(* IEC 61131-3 sources: stdmachine/plc/src/03_Base, 34 files *)

(* ---- GVL_BeaconBits.st ---- *)
// Codage de la balise (ST_MachineStatus.nBeacon, ST_StationStatus.nBeacon, I_Beacon.SetPattern)
{attribute 'qualified_only'}
VAR_GLOBAL CONSTANT
    RED : UINT := 16#0001;
    ORANGE : UINT := 16#0002;
    GREEN : UINT := 16#0004;
    BLUE : UINT := 16#0008;
    RED_BLINK : UINT := 16#0100;
    ORANGE_BLINK : UINT := 16#0200;
    GREEN_BLINK : UINT := 16#0400;
    BLUE_BLINK : UINT := 16#0800;
    BUZZER : UINT := 16#1000;
END_VAR

(* ---- GVL_Curves.st ---- *)
// Courbes de presse (docs/05 § 9) : tampon circulaire GVL_Hmi.aCurve[1..8], dernière courbe de chaque station
// pour la trace de l'opération (ST_TraceRecord.nCurveId).
{attribute 'qualified_only'}
VAR_GLOBAL
    nNextCurveId : UDINT := 1;
    nNextSlot : USINT := 1;
    aLastCurveId : ARRAY[0..GVL_Const.MAX_STATIONS] OF UDINT;
    aLastCurveTime : ARRAY[0..GVL_Const.MAX_STATIONS] OF LINT;      // début de l'enregistrement (UTC)
END_VAR

(* ---- GVL_IoRef.st ---- *)
// Pointeurs vers l'image E/S et les pools matériels du projet de la machine (docs/04 § 6).
// GVL_IO et GVL_Hw sont dans le projet de la machine (reliés aux bornes) ; MAIN les donne ici au premier cycle :
//     GVL_IoRef.pDI := ADR(GVL_IO.aDI); … ; GVL_IoRef.pAxis := ADR(GVL_Hw.aAxis); GVL_IoRef.nAxes := …
{attribute 'qualified_only'}
VAR_GLOBAL
    pDI : POINTER TO ARRAY[0..GVL_Const.MAX_DI - 1] OF BOOL;
    pDO : POINTER TO ARRAY[0..GVL_Const.MAX_DO - 1] OF BOOL;
    pAI : POINTER TO ARRAY[0..GVL_Const.MAX_AI - 1] OF INT;
    pAO : POINTER TO ARRAY[0..GVL_Const.MAX_AO - 1] OF INT;
    pAxis : POINTER TO ARRAY[1..GVL_Const.MAX_AXES] OF AXIS_REF;   // GVL_Hw.aAxis
    nAxes : INT;                     // nombre d'axes reliés dans GVL_Hw
    // Rempli par FB_Machine au premier cycle, pour les objets Système planaire et Mover
    ipPlanar : I_PlanarDriver;
    ipMovers : I_MoverMotion;
END_VAR

(* ---- GVL_Sim.st ---- *)
// Simulation de toute la machine (docs/04 § 6.3)
{attribute 'qualified_only'}
VAR_GLOBAL
    bAllSimulated : BOOL;
    nSeed : UDINT := 16#2545F491;      // générateur pseudo-aléatoire des objets simulés (F_SimRandom)
END_VAR

(* ---- F_AddDeployError.st ---- *)
// Ajoute une erreur à la réponse de déploiement (docs/05 § 10, étape 5) ; les codes sont listés dans FB_Loader
FUNCTION F_AddDeployError : BOOL
VAR_IN_OUT
    stResp : ST_DeployResponse;
END_VAR
VAR_INPUT
    nCode : UINT;
    nStation : USINT;
    nTable : USINT;
    nInstr : INT;
    nObject : UINT;
    nDetail : UDINT;
END_VAR
F_AddDeployError := FALSE;
IF stResp.nErrors >= 32 THEN RETURN; END_IF       // les suivantes sont perdues : 32 suffisent pour corriger
stResp.nErrors := stResp.nErrors + 1;
stResp.aError[stResp.nErrors].nCode := nCode;
stResp.aError[stResp.nErrors].nStation := nStation;
stResp.aError[stResp.nErrors].nTable := nTable;
stResp.aError[stResp.nErrors].nInstr := nInstr;
stResp.aError[stResp.nErrors].nObject := nObject;
stResp.aError[stResp.nErrors].nDetail := nDetail;
F_AddDeployError := TRUE;
END_FUNCTION

(* ---- F_AddRetained.st ---- *)
// Ajoute une valeur à la liste publiée pour la sauvegarde par la HMI (docs/02 § 7.4)
FUNCTION F_AddRetained : BOOL
VAR_IN_OUT
    stOut : ST_RetainedValues;
    stItem : ST_RetainedItem;
END_VAR
F_AddRetained := FALSE;
IF stOut.nCount >= 2048 THEN RETURN; END_IF
stOut.nCount := stOut.nCount + 1;
stOut.aItem[stOut.nCount] := stItem;
F_AddRetained := TRUE;
END_FUNCTION

(* ---- F_AggregateState.st ---- *)
// État agrégé d'un parent : En erreur > Non initialisé > En cours > Prêt (docs/04 § 8)
FUNCTION F_AggregateState : E_ObjState
VAR_INPUT
    eCurrent : E_ObjState;       // agrégat en cours de calcul
    eChild : E_ObjState;
END_VAR
IF eCurrent = E_ObjState.Error OR eChild = E_ObjState.Error THEN
    F_AggregateState := E_ObjState.Error;
ELSIF eCurrent = E_ObjState.NotInitialized OR eChild = E_ObjState.NotInitialized THEN
    F_AggregateState := E_ObjState.NotInitialized;
ELSIF eCurrent = E_ObjState.Busy OR eChild = E_ObjState.Busy THEN
    F_AggregateState := E_ObjState.Busy;
ELSE
    F_AggregateState := E_ObjState.Ready;
END_IF

(* ---- F_ApplyOp.st ---- *)
// SetVar : 0 affecter, 1 ajouter, 2 soustraire (docs/06 § 3)
FUNCTION F_ApplyOp : LREAL
VAR_INPUT
    fCurrent : LREAL;
    fValue : LREAL;
    nOp : DINT;
END_VAR
CASE nOp OF
    1: F_ApplyOp := fCurrent + fValue;
    2: F_ApplyOp := fCurrent - fValue;
ELSE
    F_ApplyOp := fValue;
END_CASE

(* ---- F_AxisRef.st ---- *)
// Pointeur vers l'axe NC n° nDevice du pool matériel (docs/04 § 6.2) ; 0 si absent
FUNCTION F_AxisRef : POINTER TO AXIS_REF
VAR_INPUT
    nDevice : INT;
END_VAR
IF GVL_IoRef.pAxis = 0 OR nDevice < 1 OR nDevice > GVL_IoRef.nAxes OR nDevice > GVL_Const.MAX_AXES THEN
    F_AxisRef := 0;
ELSE
    F_AxisRef := ADR(GVL_IoRef.pAxis^[nDevice]);
END_IF

(* ---- F_BeaconPattern.st ---- *)
// Couleurs de la balise selon l'état (docs/02 § 8, tableau des balises)
FUNCTION F_BeaconPattern : UINT
VAR_INPUT
    eState : E_State;
    bMaintenance : BOOL;         // mode Maintenance, ou état déclaré maintenance, essais, nettoyage
    bOperatorAwaited : BOOL;     // mover à vider, fin d'OF, machine vidée, réaction qualité…
    bStationAborted : BOOL;      // machine : une station Aborted pendant que la machine produit
END_VAR
VAR
    n : UINT;
END_VAR
CASE eState OF
    E_State.Execute:
        n := GVL_BeaconBits.GREEN;
        IF bStationAborted THEN n := n OR GVL_BeaconBits.RED_BLINK; END_IF
    E_State.Idle:
        n := GVL_BeaconBits.GREEN_BLINK;
    E_State.Held, E_State.Stopped:
        n := GVL_BeaconBits.ORANGE;
    E_State.Resetting, E_State.Stopping, E_State.Clearing:
        n := GVL_BeaconBits.ORANGE_BLINK;
    E_State.Aborted:
        n := GVL_BeaconBits.RED_BLINK OR GVL_BeaconBits.BUZZER;
END_CASE
IF bMaintenance THEN n := n OR GVL_BeaconBits.BLUE; END_IF
IF bOperatorAwaited THEN n := n OR GVL_BeaconBits.BLUE_BLINK; END_IF
F_BeaconPattern := n;

(* ---- F_CalibStateNum.st ---- *)
// État de calibration ↔ nombre, pour la sauvegarde des valeurs par la HMI (ST_RetainedItem.aValue[1])
FUNCTION F_CalibStateNum : LREAL
VAR_INPUT
    eState : E_CalibState;
END_VAR
CASE eState OF
    E_CalibState.Valid: F_CalibStateNum := 1;
    E_CalibState.Expired: F_CalibStateNum := 2;
    E_CalibState.Failed: F_CalibStateNum := 3;
    E_CalibState.Running: F_CalibStateNum := 4;
ELSE
    F_CalibStateNum := 0;
END_CASE
END_FUNCTION

(* ---- F_CalibStateOf.st ---- *)
// Nombre → état de calibration (restauration) ; une calibration en cours à la sauvegarde revient « jamais faite »
FUNCTION F_CalibStateOf : E_CalibState
VAR_INPUT
    fValue : LREAL;
END_VAR
IF fValue > 2.5 AND fValue < 3.5 THEN
    F_CalibStateOf := E_CalibState.Failed;
ELSIF fValue > 1.5 AND fValue < 2.5 THEN
    F_CalibStateOf := E_CalibState.Expired;
ELSIF fValue > 0.5 AND fValue < 1.5 THEN
    F_CalibStateOf := E_CalibState.Valid;
ELSE
    F_CalibStateOf := E_CalibState.Never;
END_IF
END_FUNCTION

(* ---- F_CatalogBit.st ---- *)
// Vrai si le bit de l'action est posé dans un masque du catalogue (GVL_Catalog.a*Mask)
FUNCTION F_CatalogBit : BOOL
VAR_INPUT
    nMask : UDINT;
    nAction : UINT;
END_VAR
IF nAction < 1 OR nAction > GVL_Const.MAX_ACTION THEN
    F_CatalogBit := FALSE;
ELSE
    F_CatalogBit := (SHR(nMask, nAction - 1) AND 1) = 1;
END_IF

(* ---- F_CatalogHasAction.st ---- *)
// L'action existe-t-elle pour ce type ? (docs/04 § 7.3)
FUNCTION F_CatalogHasAction : BOOL
VAR_INPUT
    nType : UINT;
    nAction : UINT;
END_VAR
IF nType > GVL_Const.MAX_TYPE THEN
    F_CatalogHasAction := FALSE;
ELSE
    F_CatalogHasAction := F_CatalogBit(GVL_Catalog.aActionMask[nType], nAction);
END_IF

(* ---- F_Compare.st ---- *)
// Terme de condition (docs/05 § 3.7) : égalités sur réels à 1e-9 près
FUNCTION F_Compare : BOOL
VAR_INPUT
    a : LREAL;
    eCmp : E_Cmp;
    b : LREAL;
END_VAR
CASE eCmp OF
    E_Cmp.Eq: F_Compare := ABS(a - b) < 1.0E-9;
    E_Cmp.Ne: F_Compare := ABS(a - b) >= 1.0E-9;
    E_Cmp.Lt: F_Compare := a < b;
    E_Cmp.Le: F_Compare := a <= b + 1.0E-9;
    E_Cmp.Gt: F_Compare := a > b;
    E_Cmp.Ge: F_Compare := a >= b - 1.0E-9;
    E_Cmp.IsTrue: F_Compare := a <> 0;
    E_Cmp.IsFalse: F_Compare := a = 0;
ELSE
    F_Compare := FALSE;
END_CASE

(* ---- F_CycleMs.st ---- *)
// Durée du cycle de la tâche courante en ms (docs/04 § 2)
FUNCTION F_CycleMs : LREAL
VAR
    nTask : DINT;
END_VAR
nTask := GETCURTASKINDEXEX();
F_CycleMs := UDINT_TO_LREAL(TwinCAT_SystemInfoVarList._TaskInfo[nTask].CycleTime) / 10000.0;

(* ---- F_Pad.st ---- *)
// Nombre écrit sur nWidth chiffres, complété par des zéros
FUNCTION F_Pad : STRING(10)
VAR_INPUT
    nValue : UDINT;
    nWidth : INT;
END_VAR
F_Pad := UDINT_TO_STRING(nValue);
WHILE LEN(F_Pad) < nWidth DO
    F_Pad := CONCAT('0', F_Pad);
END_WHILE

(* ---- F_ParamSpeed.st ---- *)
// Vitesse d'un paramètre résolu, en % de la Vmax (docs/04 § 12) : n° de vitesse V1..V8 ou % direct
FUNCTION F_ParamSpeed : LREAL
VAR_INPUT
    refParams : REFERENCE TO ST_ActParams;
    nParam : USINT;
    refCfg : REFERENCE TO ST_ObjConfig;
    nDefaultSpeed : USINT;       // V utilisé si le paramètre est absent
END_VAR
VAR
    nV : INT;
END_VAR
IF nParam >= 1 AND nParam <= GVL_Const.MAX_PARAMS THEN
    CASE refParams.aKind[nParam] OF
        E_ParamKind.SpeedPercent:
            F_ParamSpeed := LIMIT(0.0, refParams.aReal[nParam], 100.0);
            RETURN;
        E_ParamKind.SpeedIndex, E_ParamKind.Real:
            nV := LREAL_TO_INT(refParams.aReal[nParam]);
            IF nV >= 1 AND nV <= GVL_Const.MAX_SPEEDS AND refCfg.aSpeedPct[nV] > 0 THEN
                F_ParamSpeed := refCfg.aSpeedPct[nV];
                RETURN;
            END_IF
    END_CASE
END_IF
IF nDefaultSpeed >= 1 AND nDefaultSpeed <= GVL_Const.MAX_SPEEDS AND refCfg.aSpeedPct[nDefaultSpeed] > 0 THEN
    F_ParamSpeed := refCfg.aSpeedPct[nDefaultSpeed];
ELSE
    F_ParamSpeed := 50.0;
END_IF

(* ---- F_PartId.st ---- *)
// Identifiant de pièce généré (docs/05 § 5.5) : <machine>-<AAAAMMJJ>-<compteur sur 6 chiffres>
FUNCTION F_PartId : STRING(40)
VAR_INPUT
    sMachine : STRING(40);
    nCounter : UDINT;
END_VAR
VAR
    stFt : T_FILETIME;
    stTime : TIMESTRUCT;
    nNow : ULINT;
    sDate : STRING(10);
    sNum : STRING(10);
END_VAR
nNow := F_GetSystemTime();
stFt.dwLowDateTime := ULINT_TO_DWORD(nNow AND 16#FFFFFFFF);
stFt.dwHighDateTime := ULINT_TO_DWORD(SHR(nNow, 32));
stTime := FILETIME_TO_SYSTEMTIME(stFt);
sDate := CONCAT(WORD_TO_STRING(stTime.wYear), CONCAT(F_Pad(WORD_TO_UDINT(stTime.wMonth), 2), F_Pad(WORD_TO_UDINT(stTime.wDay), 2)));
sNum := F_Pad(nCounter MOD 1000000, 6);
F_PartId := CONCAT(CONCAT(CONCAT(sMachine, '-'), sDate), CONCAT('-', sNum));

(* ---- F_ReadAI.st ---- *)
// Lecture brute d'une entrée analogique (docs/04 § 6.1) : référence invalide -> 0
FUNCTION F_ReadAI : INT
VAR_INPUT
    stRef : ST_SignalRef;
END_VAR
IF stRef.eKind <> E_SignalKind.AI OR GVL_IoRef.pAI = 0 OR stRef.nIndex < 0 OR stRef.nIndex >= GVL_Const.MAX_AI THEN
    F_ReadAI := 0;
    RETURN;
END_IF
F_ReadAI := GVL_IoRef.pAI^[stRef.nIndex];

(* ---- F_ReadDI.st ---- *)
// Lecture d'une entrée numérique par référence (docs/04 § 6.1) : référence invalide -> FALSE
FUNCTION F_ReadDI : BOOL
VAR_INPUT
    stRef : ST_SignalRef;
END_VAR
IF stRef.eKind <> E_SignalKind.DI OR GVL_IoRef.pDI = 0 OR stRef.nIndex < 0 OR stRef.nIndex >= GVL_Const.MAX_DI THEN
    F_ReadDI := FALSE;
    RETURN;
END_IF
F_ReadDI := GVL_IoRef.pDI^[stRef.nIndex] XOR stRef.bInvert;

(* ---- F_SignalValid.st ---- *)
// Vrai si la référence désigne un signal du bon type dans l'image E/S
FUNCTION F_SignalValid : BOOL
VAR_INPUT
    stRef : ST_SignalRef;
    eKind : E_SignalKind;
END_VAR
F_SignalValid := stRef.eKind = eKind AND stRef.nIndex >= 0;

(* ---- F_SimRandom.st ---- *)
// Nombre pseudo-aléatoire dans [0, 1) pour les objets simulés (générateur congruentiel, Numerical Recipes)
FUNCTION F_SimRandom : LREAL
GVL_Sim.nSeed := GVL_Sim.nSeed * 1664525 + 1013904223;
F_SimRandom := UDINT_TO_LREAL(GVL_Sim.nSeed) / 4294967296.0;
END_FUNCTION

(* ---- F_StartRefusalCode.st ---- *)
// Code d'erreur commune correspondant au refus d'un Start (docs/03 § 1.3)
FUNCTION F_StartRefusalCode : UINT
VAR_INPUT
    eStart : E_StartResult;
END_VAR
CASE eStart OF
    E_StartResult.Busy, E_StartResult.NotReady: F_StartRefusalCode := GVL_Catalog.Err_NotReady;
    E_StartResult.UnknownAction: F_StartRefusalCode := GVL_Catalog.Err_UnknownAction;
    E_StartResult.BadParam: F_StartRefusalCode := GVL_Catalog.Err_BadParam;
    E_StartResult.Interlocked: F_StartRefusalCode := GVL_Catalog.Err_Interlocked;
    E_StartResult.Disabled: F_StartRefusalCode := GVL_Catalog.Err_Disabled;
    E_StartResult.ManualOnly: F_StartRefusalCode := GVL_Catalog.Err_ManualOnly;
    E_StartResult.NotConfigured: F_StartRefusalCode := GVL_Catalog.Err_NotWired;
ELSE
    F_StartRefusalCode := GVL_Catalog.Err_NotReady;
END_CASE

(* ---- F_Verdict.st ---- *)
// Verdict d'une pièce depuis sa donnée 1 (0 non défini, 1 bon, 2 mauvais)
FUNCTION F_Verdict : E_Verdict
VAR_INPUT
    fData : LREAL;
END_VAR
IF fData > 1.5 THEN
    F_Verdict := E_Verdict.Bad;
ELSIF fData > 0.5 THEN
    F_Verdict := E_Verdict.Good;
ELSE
    F_Verdict := E_Verdict.Undefined;
END_IF
END_FUNCTION

(* ---- F_WriteAO.st ---- *)
// Écriture brute d'une sortie analogique (docs/04 § 6.1) : référence invalide -> ignorée
FUNCTION F_WriteAO : BOOL
VAR_INPUT
    stRef : ST_SignalRef;
    nValue : INT;
END_VAR
IF stRef.eKind <> E_SignalKind.AO OR GVL_IoRef.pAO = 0 OR stRef.nIndex < 0 OR stRef.nIndex >= GVL_Const.MAX_AO THEN
    F_WriteAO := FALSE;
    RETURN;
END_IF
GVL_IoRef.pAO^[stRef.nIndex] := nValue;
F_WriteAO := TRUE;

(* ---- F_WriteDO.st ---- *)
// Écriture d'une sortie numérique par référence (docs/04 § 6.1) : référence invalide -> ignorée
FUNCTION F_WriteDO : BOOL
VAR_INPUT
    stRef : ST_SignalRef;
    bValue : BOOL;
END_VAR
IF stRef.eKind <> E_SignalKind.DO OR GVL_IoRef.pDO = 0 OR stRef.nIndex < 0 OR stRef.nIndex >= GVL_Const.MAX_DO THEN
    F_WriteDO := FALSE;
    RETURN;
END_IF
GVL_IoRef.pDO^[stRef.nIndex] := bValue XOR stRef.bInvert;
F_WriteDO := TRUE;

(* ---- FB_AlarmManager.st ---- *)
// Alarmes actives et tampon d'événements (docs/04 § 10, docs/14 § 5).
// Une alarme est identifiée par (n° global, code) ; la lever deux fois ne la duplique pas.
// Les données vivent dans GVL_Hmi.stAlarms (Bind), pour que la HMI les lise sans copie.
FUNCTION_BLOCK FB_AlarmManager IMPLEMENTS I_AlarmSink
VAR
    _refBuf : REFERENCE TO ST_AlarmBuffer;
    _stCtx : ST_AlarmContext;          // contexte de la prochaine alarme (SetContext)
    _aLatched : ARRAY[1..GVL_Const.ALARM_ACTIVE] OF BOOL;   // alarme sans cause durable : close à l'acquittement
    nLost : UDINT;                     // alarmes perdues, liste pleine
END_VAR

METHOD Bind
VAR_INPUT
    refBuf : REFERENCE TO ST_AlarmBuffer;
END_VAR
_refBuf REF= refBuf;
END_METHOD

METHOD SetContext
VAR_INPUT
    stCtx : ST_AlarmContext;
END_VAR
_stCtx := stCtx;
END_METHOD

// Alarme sur condition (erreur d'objet) : reste active jusqu'à Clear
METHOD Raise
VAR_INPUT
    nGlobalId : UDINT;
    nCode : UINT;
    nSubCode : UDINT;
    eSeverity : E_Severity;
END_VAR
_Raise(nGlobalId, nCode, nSubCode, eSeverity, FALSE);
END_METHOD

// Alarme sur événement (séquenceurs, process) : close dès qu'elle est acquittée
METHOD RaiseEvent
VAR_INPUT
    nGlobalId : UDINT;
    nCode : UINT;
    nSubCode : UDINT;
    eSeverity : E_Severity;
END_VAR
_Raise(nGlobalId, nCode, nSubCode, eSeverity, TRUE);
END_METHOD

// La cause a disparu
METHOD Clear
VAR_INPUT
    nGlobalId : UDINT;
    nCode : UINT;
END_VAR
VAR
    i : INT;
END_VAR
IF NOT __ISVALIDREF(_refBuf) THEN RETURN; END_IF
i := _Find(nGlobalId, nCode);
IF i = 0 THEN RETURN; END_IF
IF _refBuf.aActive[i].eState = E_AlarmState.ActiveUnacked THEN
    _refBuf.aActive[i].eState := E_AlarmState.ClearedUnacked;
    _refBuf.aActive[i].tCleared := F_NowUtc();
    _Event(E_AlarmEvent.Cleared, i, '');
ELSIF _refBuf.aActive[i].eState = E_AlarmState.ActiveAcked THEN
    _refBuf.aActive[i].tCleared := F_NowUtc();
    _Close(i, '');
END_IF
END_METHOD

// Acquittement d'un avertissement par l'opérateur (nGlobalId 0 = tous les avertissements)
METHOD AckWarning
VAR_INPUT
    nGlobalId : UDINT;
    nCode : UINT;
    sUser : STRING(24);
END_VAR
VAR
    i : INT;
END_VAR
IF NOT __ISVALIDREF(_refBuf) THEN RETURN; END_IF
i := _refBuf.nActive;
WHILE i >= 1 DO
    IF _refBuf.aActive[i].eSeverity = E_Severity.Warning
       AND (nGlobalId = 0 OR (_refBuf.aActive[i].nGlobalId = nGlobalId AND _refBuf.aActive[i].nCode = nCode)) THEN
        _Ack(i, sUser);
    END_IF
    i := i - 1;
END_WHILE
END_METHOD

// Acquittement des défauts d'une station (Clearing) ou de la machine (nStation 0 : toutes les alarmes de défaut)
METHOD AckFaults
VAR_INPUT
    nStation : UINT;
    bAll : BOOL;                     // machine : défauts de toutes les stations aussi
    sUser : STRING(24);
END_VAR
VAR
    i : INT;
    nSt : UINT;
END_VAR
IF NOT __ISVALIDREF(_refBuf) THEN RETURN; END_IF
i := _refBuf.nActive;
WHILE i >= 1 DO
    nSt := UDINT_TO_UINT(_refBuf.aActive[i].nGlobalId / 1000);
    IF (_refBuf.aActive[i].eSeverity = E_Severity.StationFault OR _refBuf.aActive[i].eSeverity = E_Severity.MachineFault)
       AND (bAll OR nSt = nStation) THEN
        _Ack(i, sUser);
    END_IF
    i := i - 1;
END_WHILE
END_METHOD

// Politique Refaire, Pièce mauvaise, Aller à, Ignorer : l'alarme passe en information (docs/05 § 3.6)
METHOD Downgrade
VAR_INPUT
    nGlobalId : UDINT;
    nCode : UINT;
END_VAR
VAR
    i : INT;
END_VAR
IF NOT __ISVALIDREF(_refBuf) THEN RETURN; END_IF
i := _Find(nGlobalId, nCode);
IF i = 0 THEN RETURN; END_IF
_refBuf.aActive[i].eSeverity := E_Severity.Info;
_Close(i, '');
END_METHOD

// Première alarme de défaut active d'une station (ou de la machine), pour la raison d'arrêt (docs/14 § 4)
METHOD FirstFault : INT
VAR_INPUT
    nStation : UINT;
    bAnyStation : BOOL;
END_VAR
VAR
    i : INT;
    tBest : LINT;
END_VAR
FirstFault := 0;
IF NOT __ISVALIDREF(_refBuf) THEN RETURN; END_IF
FOR i := 1 TO _refBuf.nActive DO
    IF (_refBuf.aActive[i].eSeverity = E_Severity.StationFault OR _refBuf.aActive[i].eSeverity = E_Severity.MachineFault
        OR _refBuf.aActive[i].eSeverity = E_Severity.Quality)
       AND (bAnyStation OR UDINT_TO_UINT(_refBuf.aActive[i].nGlobalId / 1000) = nStation)
       AND (FirstFault = 0 OR _refBuf.aActive[i].tRaised < tBest) THEN
        FirstFault := i;
        tBest := _refBuf.aActive[i].tRaised;
    END_IF
END_FOR
END_METHOD

METHOD MarkCause
VAR_INPUT
    nIndex : INT;
END_VAR
IF __ISVALIDREF(_refBuf) AND nIndex >= 1 AND nIndex <= _refBuf.nActive THEN _refBuf.aActive[nIndex].bCause := TRUE; END_IF
END_METHOD

// ---------- interne

METHOD PRIVATE _Raise
VAR_INPUT
    nGlobalId : UDINT;
    nCode : UINT;
    nSubCode : UDINT;
    eSeverity : E_Severity;
    bLatched : BOOL;
END_VAR
VAR
    i : INT;
END_VAR
IF NOT __ISVALIDREF(_refBuf) THEN RETURN; END_IF
i := _Find(nGlobalId, nCode);
IF i > 0 THEN
    _refBuf.aActive[i].nSubCode := nSubCode;
    _refBuf.aActive[i].nRepeat := _refBuf.aActive[i].nRepeat + 1;
    IF _refBuf.aActive[i].eState = E_AlarmState.ClearedUnacked THEN _refBuf.aActive[i].eState := E_AlarmState.ActiveUnacked; END_IF
    _Event(E_AlarmEvent.Repeated, i, '');
    RETURN;
END_IF
IF _refBuf.nActive >= GVL_Const.ALARM_ACTIVE THEN
    nLost := nLost + 1;
    RETURN;
END_IF
_refBuf.nActive := _refBuf.nActive + 1;
i := _refBuf.nActive;
_refBuf.aActive[i].nGlobalId := nGlobalId;
_refBuf.aActive[i].nCode := nCode;
_refBuf.aActive[i].nSubCode := nSubCode;
_refBuf.aActive[i].eSeverity := eSeverity;
_refBuf.aActive[i].eState := E_AlarmState.ActiveUnacked;
_refBuf.aActive[i].tRaised := F_NowUtc();
_refBuf.aActive[i].tCleared := 0;
_refBuf.aActive[i].nRepeat := 0;
_refBuf.aActive[i].bCause := FALSE;
_refBuf.aActive[i].stCtx := _stCtx;
_aLatched[i] := bLatched;
_Event(E_AlarmEvent.Raised, i, '');
MEMSET(ADR(_stCtx), 0, SIZEOF(_stCtx));
IF eSeverity = E_Severity.Info THEN _Close(i, ''); END_IF    // une information est close dès son apparition
END_METHOD

METHOD PRIVATE _Ack
VAR_INPUT
    i : INT;
    sUser : STRING(24);
END_VAR
CASE _refBuf.aActive[i].eState OF
    E_AlarmState.ActiveUnacked:
        IF _aLatched[i] THEN
            _Close(i, sUser);
        ELSE
            _refBuf.aActive[i].eState := E_AlarmState.ActiveAcked;
            _Event(E_AlarmEvent.Acked, i, sUser);
        END_IF
    E_AlarmState.ClearedUnacked:
        _Close(i, sUser);
END_CASE
END_METHOD

METHOD PRIVATE _Close
VAR_INPUT
    i : INT;
    sUser : STRING(24);
END_VAR
VAR
    k : INT;
END_VAR
_Event(E_AlarmEvent.Closed, i, sUser);
FOR k := i TO _refBuf.nActive - 1 DO
    _refBuf.aActive[k] := _refBuf.aActive[k + 1];
    _aLatched[k] := _aLatched[k + 1];
END_FOR
MEMSET(ADR(_refBuf.aActive[_refBuf.nActive]), 0, SIZEOF(_refBuf.aActive[1]));
_aLatched[_refBuf.nActive] := FALSE;
_refBuf.nActive := _refBuf.nActive - 1;
END_METHOD

METHOD PRIVATE _Find : INT
VAR_INPUT
    nGlobalId : UDINT;
    nCode : UINT;
END_VAR
VAR
    i : INT;
END_VAR
_Find := 0;
FOR i := 1 TO _refBuf.nActive DO
    IF _refBuf.aActive[i].nGlobalId = nGlobalId AND _refBuf.aActive[i].nCode = nCode THEN
        _Find := i;
        RETURN;
    END_IF
END_FOR
END_METHOD

METHOD PRIVATE _Event
VAR_INPUT
    eEvent : E_AlarmEvent;
    i : INT;
    sUser : STRING(24);
END_VAR
VAR
    k : INT;
END_VAR
_refBuf.nWriteSeq := _refBuf.nWriteSeq + 1;
k := UDINT_TO_INT(_refBuf.nWriteSeq MOD INT_TO_UDINT(GVL_Const.ALARM_EVENTS));
_refBuf.aEvent[k].nSeq := _refBuf.nWriteSeq;
_refBuf.aEvent[k].eEvent := eEvent;
_refBuf.aEvent[k].tTime := F_NowUtc();
_refBuf.aEvent[k].stAlarm := _refBuf.aActive[i];
_refBuf.aEvent[k].sUser := sUser;
END_METHOD
END_FUNCTION_BLOCK

(* ---- FB_Crc32.st ---- *)
// CRC-32 IEEE 802.3 (polynôme réfléchi 16#EDB88320, init et xor final 16#FFFFFFFF), calculé par tranches pour
// ne pas dépasser le temps de cycle (docs/06 § 1). Même résultat que System.IO.Hashing.Crc32 côté HMI.
FUNCTION_BLOCK FB_Crc32
VAR
    _aTable : ARRAY[0..255] OF DWORD;
    _bTable : BOOL;
    _pData : POINTER TO BYTE;
    _nSize : UDINT;
    _nDone : UDINT;
    _nCrc : DWORD;
END_VAR

METHOD Begin
VAR_INPUT
    pData : POINTER TO BYTE;
    nSize : UDINT;
END_VAR
VAR
    i : UINT;
    k : USINT;
    c : DWORD;
END_VAR
IF NOT _bTable THEN
    FOR i := 0 TO 255 DO
        c := UINT_TO_DWORD(i);
        FOR k := 1 TO 8 DO
            IF (c AND 1) = 1 THEN c := SHR(c, 1) XOR 16#EDB88320; ELSE c := SHR(c, 1); END_IF
        END_FOR
        _aTable[i] := c;
    END_FOR
    _bTable := TRUE;
END_IF
_pData := pData;
_nSize := nSize;
_nDone := 0;
_nCrc := 16#FFFFFFFF;
END_METHOD

// Traite au plus nBudget octets ; TRUE quand tout est calculé
METHOD Step : BOOL
VAR_INPUT
    nBudget : UDINT;
END_VAR
VAR
    nEnd : UDINT;
    p : POINTER TO BYTE;
END_VAR
nEnd := MIN(_nSize, _nDone + nBudget);
p := _pData + _nDone;
WHILE _nDone < nEnd DO
    _nCrc := _aTable[DWORD_TO_USINT((_nCrc XOR BYTE_TO_DWORD(p^)) AND 16#FF)] XOR SHR(_nCrc, 8);
    p := p + 1;
    _nDone := _nDone + 1;
END_WHILE
Step := _nDone >= _nSize;
END_METHOD

PROPERTY Value : UDINT
GET
Value := DWORD_TO_UDINT(_nCrc XOR 16#FFFFFFFF);
END_GET
END_PROPERTY
END_FUNCTION_BLOCK

(* ---- FB_DefaultPools.st ---- *)
// Pools d'objets par défaut de la bibliothèque (docs/04 § 9). Un projet qui a besoin d'autres tailles écrit
// son propre bloc qui implémente I_ObjectPools et le donne à FB_Machine.SetPools.
// Les axes linéaires et rotatifs partagent un pool ; tous les modules (types 100 et plus) partagent celui des groupes.
FUNCTION_BLOCK FB_DefaultPools IMPLEMENTS I_ObjectPools
VAR CONSTANT
    N_DI : UINT := 256;
    N_DO : UINT := 256;
    N_AI : UINT := 32;
    N_AO : UINT := 32;
    N_CYLINDER : UINT := 64;
    N_AXIS : UINT := 64;
    N_PLANAR : UINT := 1;
    N_MOVER : UINT := GVL_Const.MAX_MOVERS;
    N_VACUUM : UINT := 32;
    N_GRIPPER : UINT := 16;
    N_KEYENCE_IV : UINT := 8;
    N_KEYENCE_GT2 : UINT := 8;
    N_SCALE : UINT := 4;
    N_LIGHT : UINT := 16;
    N_PRESS : UINT := 8;
    N_MAGAZINE : UINT := 8;
    N_BEACON : UINT := 17;
    N_SAFETY : UINT := 17;
    N_TIMER : UINT := 32;
    N_COUNTER : UINT := 32;
    N_GROUP : UINT := 64;
END_VAR
VAR
    aDigitalInput : ARRAY[1..N_DI] OF FB_DigitalInput;
    aDigitalOutput : ARRAY[1..N_DO] OF FB_DigitalOutput;
    aAnalogInput : ARRAY[1..N_AI] OF FB_AnalogInput;
    aAnalogOutput : ARRAY[1..N_AO] OF FB_AnalogOutput;
    aCylinder : ARRAY[1..N_CYLINDER] OF FB_Cylinder;
    aAxis : ARRAY[1..N_AXIS] OF FB_Axis;
    aPlanar : ARRAY[1..N_PLANAR] OF FB_PlanarSystem;
    aMover : ARRAY[1..N_MOVER] OF FB_PlanarMover;
    aVacuum : ARRAY[1..N_VACUUM] OF FB_VacuumBlow;
    aGripper : ARRAY[1..N_GRIPPER] OF FB_Gripper;
    aKeyenceIV : ARRAY[1..N_KEYENCE_IV] OF FB_KeyenceIV;
    aKeyenceGT2 : ARRAY[1..N_KEYENCE_GT2] OF FB_KeyenceGT2;
    aScale : ARRAY[1..N_SCALE] OF FB_Scale;
    aLight : ARRAY[1..N_LIGHT] OF FB_Light;
    aPress : ARRAY[1..N_PRESS] OF FB_Press;
    aMagazine : ARRAY[1..N_MAGAZINE] OF FB_Magazine;
    aBeacon : ARRAY[1..N_BEACON] OF FB_Beacon;
    aSafety : ARRAY[1..N_SAFETY] OF FB_Safety;
    aTimer : ARRAY[1..N_TIMER] OF FB_Timer;
    aCounter : ARRAY[1..N_COUNTER] OF FB_Counter;
    aGroup : ARRAY[1..N_GROUP] OF FB_Group;
END_VAR

METHOD PoolId : UINT
VAR_INPUT
    nType : UINT;
END_VAR
IF nType = GVL_Catalog.Type_RotaryAxis THEN
    PoolId := GVL_Catalog.Type_LinearAxis;
ELSIF nType >= GVL_Catalog.Type_Group THEN
    PoolId := GVL_Catalog.Type_Group;
ELSE
    PoolId := nType;
END_IF
END_METHOD

METHOD PoolSize : UINT
VAR_INPUT
    nType : UINT;
END_VAR
CASE PoolId(nType) OF
    GVL_Catalog.Type_DigitalInput: PoolSize := N_DI;
    GVL_Catalog.Type_DigitalOutput: PoolSize := N_DO;
    GVL_Catalog.Type_AnalogInput: PoolSize := N_AI;
    GVL_Catalog.Type_AnalogOutput: PoolSize := N_AO;
    GVL_Catalog.Type_Cylinder: PoolSize := N_CYLINDER;
    GVL_Catalog.Type_LinearAxis: PoolSize := N_AXIS;
    GVL_Catalog.Type_PlanarSystem: PoolSize := N_PLANAR;
    GVL_Catalog.Type_PlanarMover: PoolSize := N_MOVER;
    GVL_Catalog.Type_VacuumBlow: PoolSize := N_VACUUM;
    GVL_Catalog.Type_Gripper: PoolSize := N_GRIPPER;
    GVL_Catalog.Type_KeyenceIV: PoolSize := N_KEYENCE_IV;
    GVL_Catalog.Type_KeyenceGT2: PoolSize := N_KEYENCE_GT2;
    GVL_Catalog.Type_Scale: PoolSize := N_SCALE;
    GVL_Catalog.Type_Light: PoolSize := N_LIGHT;
    GVL_Catalog.Type_Press: PoolSize := N_PRESS;
    GVL_Catalog.Type_Magazine: PoolSize := N_MAGAZINE;
    GVL_Catalog.Type_Beacon: PoolSize := N_BEACON;
    GVL_Catalog.Type_Safety: PoolSize := N_SAFETY;
    GVL_Catalog.Type_Timer: PoolSize := N_TIMER;
    GVL_Catalog.Type_Counter: PoolSize := N_COUNTER;
    GVL_Catalog.Type_Group: PoolSize := N_GROUP;
ELSE
    PoolSize := 0;                  // type pas encore écrit dans la bibliothèque
END_CASE
END_METHOD

METHOD Element : I_Object
VAR_INPUT
    nType : UINT;
    nIndex : UINT;
END_VAR
Element := 0;
IF nIndex < 1 OR nIndex > PoolSize(nType) THEN RETURN; END_IF
CASE PoolId(nType) OF
    GVL_Catalog.Type_DigitalInput: Element := aDigitalInput[nIndex];
    GVL_Catalog.Type_DigitalOutput: Element := aDigitalOutput[nIndex];
    GVL_Catalog.Type_AnalogInput: Element := aAnalogInput[nIndex];
    GVL_Catalog.Type_AnalogOutput: Element := aAnalogOutput[nIndex];
    GVL_Catalog.Type_Cylinder: Element := aCylinder[nIndex];
    GVL_Catalog.Type_LinearAxis: Element := aAxis[nIndex];
    GVL_Catalog.Type_PlanarSystem: Element := aPlanar[nIndex];
    GVL_Catalog.Type_PlanarMover: Element := aMover[nIndex];
    GVL_Catalog.Type_VacuumBlow: Element := aVacuum[nIndex];
    GVL_Catalog.Type_Gripper: Element := aGripper[nIndex];
    GVL_Catalog.Type_KeyenceIV: Element := aKeyenceIV[nIndex];
    GVL_Catalog.Type_KeyenceGT2: Element := aKeyenceGT2[nIndex];
    GVL_Catalog.Type_Scale: Element := aScale[nIndex];
    GVL_Catalog.Type_Light: Element := aLight[nIndex];
    GVL_Catalog.Type_Press: Element := aPress[nIndex];
    GVL_Catalog.Type_Magazine: Element := aMagazine[nIndex];
    GVL_Catalog.Type_Beacon: Element := aBeacon[nIndex];
    GVL_Catalog.Type_Safety: Element := aSafety[nIndex];
    GVL_Catalog.Type_Timer: Element := aTimer[nIndex];
    GVL_Catalog.Type_Counter: Element := aCounter[nIndex];
    GVL_Catalog.Type_Group: Element := aGroup[nIndex];
END_CASE
END_METHOD
END_FUNCTION_BLOCK

(* ---- FB_NodeBase.st ---- *)
// Nœud qui porte un override et un état agrégé : machine, station (docs/04 § 8)
FUNCTION_BLOCK FB_NodeBase IMPLEMENTS I_Node
VAR
    _ipParent : I_Node;
    _fOverride : LREAL := 100.0;    // override propre du nœud
    _fEffOverride : LREAL := 100.0;
    _eState : E_ObjState := E_ObjState.Ready;
END_VAR

METHOD SetParent
VAR_INPUT
    ipParent : I_Node;
END_VAR
_ipParent := ipParent;
END_METHOD

METHOD SetOverride
VAR_INPUT
    fPercent : LREAL;
END_VAR
_fOverride := LIMIT(0.0, fPercent, 100.0);
END_METHOD

METHOD UpdateOverride
VAR
    fParent : LREAL := 100.0;
END_VAR
IF _ipParent <> 0 THEN fParent := _ipParent.EffectiveOverride; END_IF
_fEffOverride := fParent * _fOverride / 100.0;
END_METHOD

METHOD SetState
VAR_INPUT
    eState : E_ObjState;
END_VAR
_eState := eState;
END_METHOD

PROPERTY EffectiveOverride : LREAL
GET
EffectiveOverride := _fEffOverride;
END_GET
END_PROPERTY

PROPERTY NodeState : E_ObjState
GET
NodeState := _eState;
END_GET
END_PROPERTY

PROPERTY OwnOverride : LREAL
GET
OwnOverride := _fOverride;
END_GET
END_PROPERTY
END_FUNCTION_BLOCK

(* ---- FB_ObjectBase.st ---- *)
// Base de tous les objets élémentaires (docs/04 § 7) : identité, contrat d'action, timeout recalculé par
// l'override, verrouillages, simulation, alarmes, compteurs de maintenance, publication de l'état.
// Les types dérivés redéfinissent les méthodes protégées « _… » ; les valeurs par défaut viennent du catalogue.
FUNCTION_BLOCK FB_ObjectBase IMPLEMENTS I_Object, I_Maintained
VAR
    _stInfo : ST_ObjectInfo;
    _refCfg : REFERENCE TO ST_ObjConfig;
    _ipParent : I_Node;
    _ipLocks : I_InterlockProvider;
    _ipAlarms : I_AlarmSink;
    _eState : E_ObjState := E_ObjState.NotInitialized;
    _eActStatus : E_ActStatus := E_ActStatus.Idle;
    _nAction : UINT;
    _stParams : ST_ActParams;
    _stResults : ST_ActResults;
    _stStatus : ST_ObjStatus;
    _bManual : BOOL;
    _fProgressMs : LREAL;           // temps d'action compté au prorata de l'override (actions de mouvement)
    _nTimeoutMs : UDINT;
    _fElapsedMs : LREAL;            // durée réelle de l'action
    _fEffOverride : LREAL := 100.0;
    _nErrorCode : UINT;
    _nSubCode : UDINT;
    _bInitialized : BOOL;           // posé par le type dérivé à la fin de son Init
    _eFaultSeverity : E_Severity := E_Severity.StationFault;
    _aForced : ARRAY[1..GVL_Const.MAX_SIGNALS] OF BOOL;     // simulation : entrée forcée par la HMI
    _aForcedValue : ARRAY[1..GVL_Const.MAX_SIGNALS] OF LREAL;
    _bNewObject : BOOL;             // Configure : l'élément de pool change d'objet (valeurs persistantes du type à remettre à zéro)
END_VAR
VAR PERSISTENT
    _nStableId : UDINT;             // objet du projet auquel appartiennent ces compteurs (D92)
    _nActionCount : UDINT;
    _nErrorCount : UDINT;
    _fMotionHours : LREAL;
END_VAR

METHOD Configure : BOOL
VAR_INPUT
    refCfg : REFERENCE TO ST_ObjConfig;
    nStation : UINT;
    nPoolIndex : UINT;
    ipParent : I_Node;
    ipLocks : I_InterlockProvider;
    ipAlarms : I_AlarmSink;
END_VAR
_refCfg REF= refCfg;
_ipParent := ipParent;
_ipLocks := ipLocks;
_ipAlarms := ipAlarms;
_stInfo.nStation := nStation;
_stInfo.nLocalId := refCfg.nLocalId;
_stInfo.nParentId := refCfg.nParentId;
_stInfo.nType := refCfg.nType;
_stInfo.nPoolIndex := nPoolIndex;
_stInfo.nStableId := refCfg.nStableId;
_stInfo.sName := refCfg.sName;
_stInfo.nGlobalId := UINT_TO_UDINT(nStation) * 1000 + UINT_TO_UDINT(refCfg.nLocalId);
_eFaultSeverity := SEL(nStation = 0, E_Severity.StationFault, E_Severity.MachineFault);

// Un élément de pool repris par un autre objet repart de compteurs nuls (D92)
_bNewObject := _nStableId <> refCfg.nStableId;
IF _bNewObject THEN
    _nStableId := refCfg.nStableId;
    _nActionCount := 0;
    _nErrorCount := 0;
    _fMotionHours := 0;
END_IF

_eActStatus := E_ActStatus.Idle;
_nAction := 0;
_nErrorCode := 0;
_nSubCode := 0;
_bManual := FALSE;
_bInitialized := FALSE;
_fEffOverride := 100.0;
MEMSET(ADR(_aForced), 0, SIZEOF(_aForced));
MEMSET(ADR(_stResults), 0, SIZEOF(_stResults));

IF NOT _OnConfigure() THEN
    _eState := E_ObjState.Error;
    _nErrorCode := GVL_Catalog.Err_NotWired;
    Configure := FALSE;
    RETURN;
END_IF
IF refCfg.bDisabled THEN
    _eState := E_ObjState.Disabled;
ELSIF _NeedsInit() THEN
    _eState := E_ObjState.NotInitialized;
ELSE
    _eState := E_ObjState.Ready;
END_IF
Configure := TRUE;
END_METHOD

METHOD Start : E_StartResult
VAR_INPUT
    nAction : UINT;
    refParams : REFERENCE TO ST_ActParams;
    bManual : BOOL;
END_VAR
VAR
    nLock : INT;
    nCfgTimeout : UDINT;
END_VAR
IF NOT __ISVALIDREF(_refCfg) THEN Start := E_StartResult.NotConfigured; RETURN; END_IF
IF _eState = E_ObjState.Disabled THEN Start := E_StartResult.Disabled; RETURN; END_IF
IF _eState = E_ObjState.Busy THEN Start := E_StartResult.Busy; RETURN; END_IF
IF NOT F_CatalogHasAction(_stInfo.nType, nAction) THEN Start := E_StartResult.UnknownAction; RETURN; END_IF
IF _IsManualOnly(nAction) AND NOT bManual THEN Start := E_StartResult.ManualOnly; RETURN; END_IF
IF _eState = E_ObjState.Error THEN Start := E_StartResult.NotReady; RETURN; END_IF
IF _eState = E_ObjState.NotInitialized AND NOT _IsAllowedNotInit(nAction) THEN
    Start := E_StartResult.NotReady;
    RETURN;
END_IF

_stParams := refParams;
IF NOT _ValidateParams(nAction) THEN Start := E_StartResult.BadParam; RETURN; END_IF

IF _ipLocks <> 0 THEN
    nLock := _ipLocks.Check(_stInfo.nLocalId, nAction);
    IF nLock <> 0 THEN
        _stStatus.nInterlock := INT_TO_USINT(nLock);
        Start := E_StartResult.Interlocked;
        RETURN;
    END_IF
END_IF
_stStatus.nInterlock := 0;

// Acceptée
_nAction := nAction;
_bManual := bManual;
_fProgressMs := 0;
_fElapsedMs := 0;
IF nAction <= GVL_Const.MAX_ACTION_TIMEOUTS THEN nCfgTimeout := _refCfg.aTimeoutMs[nAction]; ELSE nCfgTimeout := 0; END_IF
IF _stParams.nTimeoutMs > 0 THEN
    _nTimeoutMs := _stParams.nTimeoutMs;
ELSIF nCfgTimeout > 0 THEN
    _nTimeoutMs := nCfgTimeout;
ELSE
    _nTimeoutMs := _DefaultTimeoutMs(nAction);
END_IF
MEMSET(ADR(_stResults), 0, SIZEOF(_stResults));
_nErrorCode := 0;
_nSubCode := 0;
_nActionCount := _nActionCount + 1;
_eState := E_ObjState.Busy;
_eActStatus := _OnStart(nAction);       // Busy, ou Done / Error immédiat
IF _eActStatus <> E_ActStatus.Busy THEN
    _EndAction();
END_IF
Start := E_StartResult.Accepted;
END_METHOD

METHOD Cycle
VAR
    fCycleMs : LREAL;
    fParentOv : LREAL;
    nLock : INT;
END_VAR
IF NOT __ISVALIDREF(_refCfg) THEN RETURN; END_IF
fCycleMs := F_CycleMs();

// 1. Override effectif : les parents sont appelés avant leurs enfants (docs/04 § 8)
fParentOv := 100.0;
IF _ipParent <> 0 THEN fParentOv := _ipParent.EffectiveOverride; END_IF
_fEffOverride := fParentOv * LIMIT(0.0, _refCfg.fOverride, 100.0) / 100.0;
IF _bManual AND _eState = E_ObjState.Busy THEN
    _fEffOverride := _fEffOverride * _ManualOverride() / 100.0;
END_IF
_ApplyOverride(_fEffOverride);

// 2. Entrées
IF _IsSimulated() THEN _Simulate(); ELSE _ReadHw(); END_IF

// 3. Action en cours
IF _eState = E_ObjState.Busy THEN
    _fElapsedMs := _fElapsedMs + fCycleMs;
    IF _IsMotion(_nAction) THEN
        _fProgressMs := _fProgressMs + fCycleMs * _fEffOverride / 100.0;
        _fMotionHours := _fMotionHours + fCycleMs / 3600000.0;
        IF _ipLocks <> 0 THEN
            nLock := _ipLocks.Check(_stInfo.nLocalId, _nAction);
            IF nLock <> 0 THEN
                _OnAbort(_nAction);
                _stStatus.nInterlock := INT_TO_USINT(nLock);
                _Fail(GVL_Catalog.Err_Interlocked, INT_TO_UDINT(nLock));
            END_IF
        END_IF
    ELSE
        _fProgressMs := _fProgressMs + fCycleMs;
    END_IF
    IF _eState = E_ObjState.Busy THEN
        _eActStatus := _OnCycle(_nAction);
        IF _eActStatus = E_ActStatus.Busy AND _nTimeoutMs > 0 AND _fProgressMs >= UDINT_TO_LREAL(_nTimeoutMs) THEN
            _OnAbort(_nAction);
            _Fail(GVL_Catalog.Err_Timeout, _nAction);
        ELSIF _eActStatus <> E_ActStatus.Busy THEN
            _EndAction();
        END_IF
    END_IF
END_IF

// 4. Surveillance continue
IF _eState <> E_ObjState.Disabled THEN _Monitor(); END_IF

// 5. Sorties
IF NOT _IsSimulated() THEN _WriteHw(); END_IF

// 6. Publication pour la HMI
_stStatus.eState := _eState;
_stStatus.eActStatus := _eActStatus;
_stStatus.nAction := UINT_TO_USINT(_nAction);
_stStatus.bManual := _bManual;
_stStatus.nErrorCode := _nErrorCode;
_stStatus.nSubCode := _nSubCode;
_stStatus.fEffOverride := LREAL_TO_REAL(_fEffOverride);
_stStatus.bOverrideHalted := (_eState = E_ObjState.Busy) AND _IsMotion(_nAction) AND (_fEffOverride <= 0.0);
_stStatus.bSimulated := _IsSimulated();
_stStatus.nElapsedMs := LREAL_TO_UDINT(_fElapsedMs);
_stStatus.nTimeoutMs := _EffectiveTimeoutEstimate();
_stStatus.nActionCount := _nActionCount;
_stStatus.nErrorCount := _nErrorCount;
_stStatus.fMotionHours := LREAL_TO_REAL(_fMotionHours);
_stStatus.fProgress := -1;
_Publish();                             // aValue[1..4], fProgress
END_METHOD

METHOD Abort
IF _eState = E_ObjState.Busy THEN
    _OnAbort(_nAction);
    _eActStatus := E_ActStatus.Error;
    _nErrorCode := GVL_Catalog.Err_Aborted;     // action interrompue par Abort : pas d'alarme levée
    _nSubCode := _nAction;
    _eState := SEL(_NeedsInit() AND NOT _bInitialized, E_ObjState.Ready, E_ObjState.NotInitialized);
END_IF
_SafeState();
IF _HardwareFault() AND _eState <> E_ObjState.Disabled THEN _eState := E_ObjState.Error; END_IF
END_METHOD

METHOD Ack : BOOL
IF _eState <> E_ObjState.Error THEN
    Ack := TRUE;
    RETURN;
END_IF
IF _OnAck() THEN
    IF _ipAlarms <> 0 AND _nErrorCode <> 0 THEN _ipAlarms.Clear(_stInfo.nGlobalId, _nErrorCode); END_IF
    _nErrorCode := 0;
    _nSubCode := 0;
    _eActStatus := E_ActStatus.Idle;
    _eState := SEL(_NeedsInit() AND NOT _bInitialized, E_ObjState.Ready, E_ObjState.NotInitialized);
    Ack := TRUE;
END_IF
END_METHOD

METHOD ForceInput
VAR_INPUT
    nSignal : USINT;
    fValue : LREAL;
END_VAR
IF nSignal = 0 THEN
    MEMSET(ADR(_aForced), 0, SIZEOF(_aForced));
ELSIF nSignal <= GVL_Const.MAX_SIGNALS THEN
    _aForced[nSignal] := TRUE;
    _aForcedValue[nSignal] := fValue;
END_IF
END_METHOD

PROPERTY EffectiveOverride : LREAL
GET
EffectiveOverride := _fEffOverride;
END_GET
END_PROPERTY

PROPERTY NodeState : E_ObjState
GET
NodeState := _eState;
END_GET
END_PROPERTY

PROPERTY Info : REFERENCE TO ST_ObjectInfo
GET
Info REF= _stInfo;
END_GET
END_PROPERTY

PROPERTY ActStatus : E_ActStatus
GET
ActStatus := _eActStatus;
END_GET
END_PROPERTY

PROPERTY Results : REFERENCE TO ST_ActResults
GET
Results REF= _stResults;
END_GET
END_PROPERTY

PROPERTY Status : REFERENCE TO ST_ObjStatus
GET
Status REF= _stStatus;
END_GET
END_PROPERTY

// ---------- Compteurs de maintenance (I_Maintained)

PROPERTY StableId : UDINT
GET
StableId := _nStableId;
END_GET
END_PROPERTY

PROPERTY ActionCount : UDINT
GET
ActionCount := _nActionCount;
END_GET
END_PROPERTY

PROPERTY ErrorCount : UDINT
GET
ErrorCount := _nErrorCount;
END_GET
END_PROPERTY

PROPERTY MotionHours : LREAL
GET
MotionHours := _fMotionHours;
END_GET
END_PROPERTY

// Restauration des valeurs sauvegardées par la HMI (docs/05 § 10, étape 6)
METHOD RestoreCounters
VAR_INPUT
    nActions : UDINT;
    nErrors : UDINT;
    fHours : LREAL;
END_VAR
_nActionCount := nActions;
_nErrorCount := nErrors;
_fMotionHours := fHours;
END_METHOD

// ---------- Fin d'action et erreurs

METHOD PROTECTED _EndAction
IF _eActStatus = E_ActStatus.Done THEN
    _eState := SEL(_NeedsInit() AND NOT _bInitialized, E_ObjState.Ready, E_ObjState.NotInitialized);
ELSIF _eActStatus = E_ActStatus.Error AND _eState <> E_ObjState.Error THEN
    _Fail(GVL_Catalog.Err_UnknownAction, _nAction);     // le type a répondu Error sans dire pourquoi
END_IF
END_METHOD

METHOD PROTECTED _Fail
VAR_INPUT
    nCode : UINT;
    nSubCode : UDINT;
END_VAR
_eActStatus := E_ActStatus.Error;
_nErrorCode := nCode;
_nSubCode := nSubCode;
_eState := E_ObjState.Error;
_nErrorCount := _nErrorCount + 1;
IF _ipAlarms <> 0 THEN _ipAlarms.Raise(_stInfo.nGlobalId, nCode, nSubCode, _eFaultSeverity); END_IF
END_METHOD

METHOD PROTECTED _SetResult
VAR_INPUT
    nIndex : USINT;
    fValue : LREAL;
END_VAR
IF nIndex >= 1 AND nIndex <= GVL_Const.MAX_PARAMS THEN
    _stResults.aReal[nIndex] := fValue;
    _stResults.nCount := MAX(_stResults.nCount, nIndex);
END_IF
END_METHOD

METHOD PROTECTED _SetJudgement
VAR_INPUT
    nIndex : USINT;
    eJudgement : E_Judgement;
END_VAR
IF nIndex >= 1 AND nIndex <= GVL_Const.MAX_PARAMS THEN
    _stResults.aJudgement[nIndex] := eJudgement;
    _stResults.aReal[nIndex] := TO_LREAL(eJudgement);
    _stResults.nCount := MAX(_stResults.nCount, nIndex);
END_IF
END_METHOD

METHOD PROTECTED _SetResultPos
VAR_INPUT
    nIndex : USINT;
    stPos : ST_Position;
END_VAR
_stResults.stPos := stPos;
_stResults.nPosIndex := nIndex;
_stResults.nCount := MAX(_stResults.nCount, nIndex);
END_METHOD

// ---------- Aides

METHOD PROTECTED _IsSimulated : BOOL
_IsSimulated := GVL_Sim.bAllSimulated OR (__ISVALIDREF(_refCfg) AND_THEN _refCfg.bSimulated);
END_METHOD

METHOD PROTECTED _Forced : BOOL
VAR_INPUT
    nSignal : USINT;
END_VAR
_Forced := nSignal >= 1 AND nSignal <= GVL_Const.MAX_SIGNALS AND_THEN _aForced[nSignal];
END_METHOD

METHOD PROTECTED _ForcedValue : LREAL
VAR_INPUT
    nSignal : USINT;
END_VAR
IF nSignal >= 1 AND nSignal <= GVL_Const.MAX_SIGNALS THEN _ForcedValue := _aForcedValue[nSignal]; END_IF
END_METHOD

METHOD PROTECTED _Param : LREAL
VAR_INPUT
    nParam : USINT;              // P1..P24
END_VAR
IF nParam >= 1 AND nParam <= GVL_Const.MAX_OBJ_PARAMS THEN _Param := _refCfg.aParam[nParam]; END_IF
END_METHOD

METHOD PROTECTED _ParamReal : LREAL
VAR_INPUT
    nParam : USINT;              // a1..a8
    fDefault : LREAL;
END_VAR
IF nParam >= 1 AND nParam <= GVL_Const.MAX_PARAMS AND_THEN _stParams.aKind[nParam] <> E_ParamKind.Unused THEN
    _ParamReal := _stParams.aReal[nParam];
ELSE
    _ParamReal := fDefault;
END_IF
END_METHOD

METHOD PROTECTED _EffectiveTimeoutEstimate : UDINT
IF _nTimeoutMs = 0 THEN
    _EffectiveTimeoutEstimate := 0;
ELSIF _IsMotion(_nAction) AND _fEffOverride <= 0.0 THEN
    _EffectiveTimeoutEstimate := 16#FFFFFFFF;          // « infini » à 0 %
ELSIF _IsMotion(_nAction) THEN
    _EffectiveTimeoutEstimate := LREAL_TO_UDINT(MIN(UDINT_TO_LREAL(_nTimeoutMs) * 100.0 / _fEffOverride, 86400000.0));
ELSE
    _EffectiveTimeoutEstimate := _nTimeoutMs;
END_IF
END_METHOD

// ---------- Méthodes à redéfinir par les types (valeurs par défaut tirées du catalogue)

METHOD PROTECTED _OnConfigure : BOOL
_OnConfigure := TRUE;
END_METHOD

METHOD PROTECTED _NeedsInit : BOOL
_NeedsInit := FALSE;
END_METHOD

METHOD PROTECTED _IsMotion : BOOL
VAR_INPUT
    nAction : UINT;
END_VAR
_IsMotion := _stInfo.nType <= GVL_Const.MAX_TYPE AND_THEN F_CatalogBit(GVL_Catalog.aMotionMask[_stInfo.nType], nAction);
END_METHOD

METHOD PROTECTED _IsAllowedNotInit : BOOL
VAR_INPUT
    nAction : UINT;
END_VAR
_IsAllowedNotInit := FALSE;
END_METHOD

METHOD PROTECTED _IsManualOnly : BOOL
VAR_INPUT
    nAction : UINT;
END_VAR
_IsManualOnly := _stInfo.nType <= GVL_Const.MAX_TYPE AND_THEN F_CatalogBit(GVL_Catalog.aManualOnlyMask[_stInfo.nType], nAction);
END_METHOD

METHOD PROTECTED _ValidateParams : BOOL
VAR_INPUT
    nAction : UINT;
END_VAR
_ValidateParams := TRUE;
END_METHOD

METHOD PROTECTED _DefaultTimeoutMs : UDINT
VAR_INPUT
    nAction : UINT;
END_VAR
IF _stInfo.nType <= GVL_Const.MAX_TYPE AND nAction >= 1 AND nAction <= GVL_Const.MAX_ACTION THEN
    _DefaultTimeoutMs := GVL_Catalog.aDefaultTimeoutMs[_stInfo.nType, nAction];
ELSE
    _DefaultTimeoutMs := 0;
END_IF
END_METHOD

METHOD PROTECTED _OnStart : E_ActStatus
VAR_INPUT
    nAction : UINT;
END_VAR
_OnStart := E_ActStatus.Error;
END_METHOD

METHOD PROTECTED _OnCycle : E_ActStatus
VAR_INPUT
    nAction : UINT;
END_VAR
_OnCycle := E_ActStatus.Done;
END_METHOD

METHOD PROTECTED _OnAbort
VAR_INPUT
    nAction : UINT;
END_VAR
;
END_METHOD

METHOD PROTECTED _SafeState
;
END_METHOD

METHOD PROTECTED _Monitor
;
END_METHOD

METHOD PROTECTED _OnAck : BOOL
_OnAck := TRUE;
END_METHOD

METHOD PROTECTED _HardwareFault : BOOL
_HardwareFault := FALSE;
END_METHOD

METHOD PROTECTED _ReadHw
;
END_METHOD

METHOD PROTECTED _WriteHw
;
END_METHOD

METHOD PROTECTED _Simulate
;
END_METHOD

METHOD PROTECTED _Publish
;
END_METHOD

METHOD PROTECTED _ApplyOverride
VAR_INPUT
    fPercent : LREAL;
END_VAR
;
END_METHOD

METHOD PROTECTED _ManualOverride : LREAL
_ManualOverride := 100.0;
END_METHOD
END_FUNCTION_BLOCK

(* ---- FB_ObjectFactory.st ---- *)
// Fabrique d'objets (docs/04 § 9) : attribue à chaque objet configuré un élément de son pool et le configure.
// Un objet déjà présent au déploiement précédent (même nStableId) reprend le même élément, pour garder ses
// compteurs de maintenance persistants (D92). Hôte 0 = la machine, 1..16 = les stations.
FUNCTION_BLOCK FB_ObjectFactory
VAR
    _ipPools : I_ObjectPools;
    _ipAlarms : I_AlarmSink;
    _aHost : ARRAY[0..GVL_Const.MAX_STATIONS] OF I_ObjectHost;
    _aNode : ARRAY[0..GVL_Const.MAX_STATIONS] OF I_Node;
    _aLocks : ARRAY[0..GVL_Const.MAX_STATIONS] OF I_InterlockProvider;
    _aUsed : ARRAY[0..GVL_Const.MAX_TYPE, 0..7] OF DWORD;    // bit = élément de pool pris par ce déploiement
    _aAssign : ARRAY[0..GVL_Const.MAX_STATIONS, 1..GVL_Const.MAX_OBJ_PER_STATION] OF UINT;  // élément attribué
END_VAR

METHOD SetPools
VAR_INPUT
    ipPools : I_ObjectPools;
    ipAlarms : I_AlarmSink;
END_VAR
_ipPools := ipPools;
_ipAlarms := ipAlarms;
END_METHOD

METHOD SetHost
VAR_INPUT
    nHost : USINT;
    ipHost : I_ObjectHost;
    ipNode : I_Node;
    ipLocks : I_InterlockProvider;
END_VAR
IF nHost <= GVL_Const.MAX_STATIONS THEN
    _aHost[nHost] := ipHost;
    _aNode[nHost] := ipNode;
    _aLocks[nHost] := ipLocks;
END_IF
END_METHOD

// Taille du pool d'un type (identité du PLC)
METHOD PoolSize : UINT
VAR_INPUT
    nType : UINT;
END_VAR
IF _ipPools <> 0 THEN PoolSize := _ipPools.PoolSize(nType); END_IF
END_METHOD

// Vérification sans effet (docs/05 § 10, étape 3) : types connus et pools suffisants pour la zone d'attente
METHOD Check : BOOL
VAR_IN_OUT
    stStaging : ST_Staging;
    stResp : ST_DeployResponse;
END_VAR
VAR
    aNeed : ARRAY[0..GVL_Const.MAX_TYPE] OF UINT;
    n : USINT;
    k : UINT;
    nCount : UINT;
    nType : UINT;
    nPool : UINT;
END_VAR
Check := TRUE;
IF _ipPools = 0 THEN
    F_AddDeployError(stResp, 7, 0, 0, 0, 0, 0);
    Check := FALSE;
    RETURN;
END_IF
FOR n := 0 TO GVL_Const.MAX_STATIONS DO
    IF n = 0 THEN nCount := stStaging.stMachine.nMachineObj; ELSE nCount := stStaging.aStation[n].nObjCount; END_IF
    FOR k := 1 TO MIN(nCount, GVL_Const.MAX_OBJ_PER_STATION) DO
        IF n = 0 THEN
            IF k > GVL_Const.MAX_MACHINE_OBJ THEN EXIT; END_IF
            nType := stStaging.stMachine.aMachineObj[k].nType;
        ELSE
            nType := stStaging.aStation[n].aObj[k].nType;
        END_IF
        IF nType = 0 OR nType > GVL_Const.MAX_TYPE OR_ELSE (GVL_Catalog.aActionMask[nType] = 0 AND nType < GVL_Catalog.Type_Group) THEN
            F_AddDeployError(stResp, 4, n, 0, 0, k, nType);         // type inconnu du catalogue du PLC
            Check := FALSE;
        ELSE
            nPool := _ipPools.PoolId(nType);
            IF nPool <= GVL_Const.MAX_TYPE THEN aNeed[nPool] := aNeed[nPool] + 1; END_IF
        END_IF
    END_FOR
END_FOR
FOR nPool := 0 TO GVL_Const.MAX_TYPE DO
    IF aNeed[nPool] > _ipPools.PoolSize(nPool) THEN
        F_AddDeployError(stResp, 7, 0, 0, 0, aNeed[nPool], nPool);  // pool trop petit (nObject = nombre demandé)
        Check := FALSE;
    END_IF
END_FOR
END_METHOD

// Attribution et configuration de tous les objets de la zone active (machine Stopped)
METHOD Build : BOOL
VAR_IN_OUT
    stResp : ST_DeployResponse;
END_VAR
VAR
    n : USINT;
    k : UINT;
    nCount : UINT;
    idx : UINT;
    pCfg : POINTER TO ST_ObjConfig;
    ipObj : I_Object;
    ipParent : I_Node;
    bOk : BOOL;
END_VAR
Build := TRUE;
IF _ipPools = 0 THEN RETURN; END_IF
MEMSET(ADR(_aUsed), 0, SIZEOF(_aUsed));
MEMSET(ADR(_aAssign), 0, SIZEOF(_aAssign));
// 1. Reprise des éléments par identifiant stable
FOR n := 0 TO GVL_Const.MAX_STATIONS DO
    nCount := _Count(n);
    FOR k := 1 TO nCount DO
        pCfg := _Cfg(n, k);
        IF pCfg^.nStableId <> 0 THEN _aAssign[n, k] := _FindByStableId(pCfg^.nType, pCfg^.nStableId); END_IF
    END_FOR
END_FOR
// 2. Les autres prennent un élément libre, de préférence jamais attribué
FOR n := 0 TO GVL_Const.MAX_STATIONS DO
    nCount := _Count(n);
    FOR k := 1 TO nCount DO
        IF _aAssign[n, k] = 0 THEN
            pCfg := _Cfg(n, k);
            _aAssign[n, k] := _FindFree(pCfg^.nType);
            IF _aAssign[n, k] = 0 THEN
                F_AddDeployError(stResp, 7, n, 0, 0, k, pCfg^.nType);
                Build := FALSE;
            END_IF
        END_IF
    END_FOR
END_FOR
IF NOT Build THEN RETURN; END_IF
// 3. Configuration, parents d'abord (la configuration est rangée parents avant enfants)
FOR n := 0 TO GVL_Const.MAX_STATIONS DO
    IF _aHost[n] <> 0 THEN
        _aHost[n].ClearObjects();
        nCount := _Count(n);
        FOR k := 1 TO nCount DO
            pCfg := _Cfg(n, k);
            idx := _aAssign[n, k];
            ipObj := _ipPools.Element(pCfg^.nType, idx);
            ipParent := _aNode[n];
            IF pCfg^.nParentId >= 1 AND pCfg^.nParentId < k THEN
                ipParent := _ipPools.Element(_Cfg(n, pCfg^.nParentId)^.nType, _aAssign[n, pCfg^.nParentId]);
            END_IF
            bOk := ipObj <> 0;
            IF bOk THEN
                bOk := ipObj.Configure(refCfg := pCfg^, nStation := n, nPoolIndex := idx, ipParent := ipParent,
                                       ipLocks := _aLocks[n], ipAlarms := _ipAlarms);
            END_IF
            IF bOk THEN
                _aHost[n].SetObject(pCfg^.nLocalId, ipObj);
            ELSE
                F_AddDeployError(stResp, 20, n, 0, 0, pCfg^.nLocalId, pCfg^.nType);   // configuration refusée par l'objet
                Build := FALSE;
            END_IF
        END_FOR
    END_IF
END_FOR
END_METHOD

METHOD PRIVATE _Count : UINT
VAR_INPUT
    n : USINT;
END_VAR
IF n = 0 THEN
    _Count := MIN(GVL_Active.stMachine.nMachineObj, GVL_Const.MAX_MACHINE_OBJ);
ELSE
    _Count := MIN(GVL_Active.aStation[n].nObjCount, GVL_Const.MAX_OBJ_PER_STATION);
END_IF
END_METHOD

METHOD PRIVATE _Cfg : POINTER TO ST_ObjConfig
VAR_INPUT
    n : USINT;
    k : UINT;
END_VAR
IF n = 0 THEN _Cfg := ADR(GVL_Active.stMachine.aMachineObj[k]); ELSE _Cfg := ADR(GVL_Active.aStation[n].aObj[k]); END_IF
END_METHOD

METHOD PRIVATE _IsUsed : BOOL
VAR_INPUT
    nPool : UINT;
    idx : UINT;
END_VAR
_IsUsed := (SHR(_aUsed[nPool, (idx - 1) / 32], (idx - 1) MOD 32) AND 1) = 1;
END_METHOD

METHOD PRIVATE _Take
VAR_INPUT
    nPool : UINT;
    idx : UINT;
END_VAR
_aUsed[nPool, (idx - 1) / 32] := _aUsed[nPool, (idx - 1) / 32] OR SHL(DWORD#1, (idx - 1) MOD 32);
END_METHOD

METHOD PRIVATE _FindByStableId : UINT
VAR_INPUT
    nType : UINT;
    nStableId : UDINT;
END_VAR
VAR
    nPool : UINT;
    idx : UINT;
    ipObj : I_Object;
    ipMaint : I_Maintained;
END_VAR
_FindByStableId := 0;
nPool := _ipPools.PoolId(nType);
IF nPool > GVL_Const.MAX_TYPE THEN RETURN; END_IF
FOR idx := 1 TO MIN(_ipPools.PoolSize(nType), 256) DO
    IF NOT _IsUsed(nPool, idx) THEN
        ipObj := _ipPools.Element(nType, idx);
        IF ipObj <> 0 AND_THEN __QUERYINTERFACE(ipObj, ipMaint) AND_THEN ipMaint.StableId = nStableId THEN
            _Take(nPool, idx);
            _FindByStableId := idx;
            RETURN;
        END_IF
    END_IF
END_FOR
END_METHOD

METHOD PRIVATE _FindFree : UINT
VAR_INPUT
    nType : UINT;
END_VAR
VAR
    nPool : UINT;
    idx : UINT;
    nAny : UINT;
    ipObj : I_Object;
    ipMaint : I_Maintained;
END_VAR
_FindFree := 0;
nPool := _ipPools.PoolId(nType);
IF nPool > GVL_Const.MAX_TYPE THEN RETURN; END_IF
FOR idx := 1 TO MIN(_ipPools.PoolSize(nType), 256) DO
    IF NOT _IsUsed(nPool, idx) THEN
        IF nAny = 0 THEN nAny := idx; END_IF
        ipObj := _ipPools.Element(nType, idx);
        IF ipObj <> 0 AND_THEN __QUERYINTERFACE(ipObj, ipMaint) AND_THEN ipMaint.StableId = 0 THEN
            _Take(nPool, idx);
            _FindFree := idx;
            RETURN;
        END_IF
    END_IF
END_FOR
IF nAny > 0 THEN
    _Take(nPool, nAny);
    _FindFree := nAny;
END_IF
END_METHOD

// Objet d'un hôte, pour la restauration des compteurs (docs/05 § 10, étape 6)
METHOD FindObject : I_Object
VAR_INPUT
    nStableId : UDINT;
END_VAR
VAR
    n : USINT;
    k : UINT;
    pCfg : POINTER TO ST_ObjConfig;
END_VAR
FindObject := 0;
IF _ipPools = 0 OR nStableId = 0 THEN RETURN; END_IF
FOR n := 0 TO GVL_Const.MAX_STATIONS DO
    FOR k := 1 TO _Count(n) DO
        pCfg := _Cfg(n, k);
        IF pCfg^.nStableId = nStableId AND _aAssign[n, k] > 0 THEN
            FindObject := _ipPools.Element(pCfg^.nType, _aAssign[n, k]);
            RETURN;
        END_IF
    END_FOR
END_FOR
END_METHOD

// Compteurs de maintenance de tous les objets attribués, ajoutés à la liste publiée pour la HMI
METHOD PublishRetained
VAR_IN_OUT
    stOut : ST_RetainedValues;
END_VAR
VAR
    n : USINT;
    k : UINT;
    pCfg : POINTER TO ST_ObjConfig;
    ipObj : I_Object;
    ipMaint : I_Maintained;
    stItem : ST_RetainedItem;
END_VAR
IF _ipPools = 0 THEN RETURN; END_IF
FOR n := 0 TO GVL_Const.MAX_STATIONS DO
    FOR k := 1 TO _Count(n) DO
        pCfg := _Cfg(n, k);
        IF _aAssign[n, k] > 0 AND pCfg^.nStableId <> 0 THEN
            ipObj := _ipPools.Element(pCfg^.nType, _aAssign[n, k]);
            IF ipObj <> 0 AND_THEN __QUERYINTERFACE(ipObj, ipMaint) THEN
                MEMSET(ADR(stItem), 0, SIZEOF(stItem));
                stItem.eKind := E_RetainedKind.ObjectCounters;
                stItem.nStation := n;
                stItem.nId := pCfg^.nStableId;
                stItem.aValue[1] := UDINT_TO_LREAL(ipMaint.ActionCount);
                stItem.aValue[2] := UDINT_TO_LREAL(ipMaint.ErrorCount);
                stItem.aValue[3] := ipMaint.MotionHours;
                F_AddRetained(stOut, stItem);
            END_IF
        END_IF
    END_FOR
END_FOR
END_METHOD

METHOD Restore : BOOL
VAR_IN_OUT
    stItem : ST_RetainedItem;
END_VAR
VAR
    ipObj : I_Object;
    ipMaint : I_Maintained;
END_VAR
Restore := FALSE;
IF stItem.eKind <> E_RetainedKind.ObjectCounters THEN RETURN; END_IF
ipObj := FindObject(stItem.nId);
IF ipObj <> 0 AND_THEN __QUERYINTERFACE(ipObj, ipMaint) THEN
    ipMaint.RestoreCounters(LREAL_TO_UDINT(stItem.aValue[1]), LREAL_TO_UDINT(stItem.aValue[2]), stItem.aValue[3]);
    Restore := TRUE;
END_IF
END_METHOD
END_FUNCTION_BLOCK

(* ---- FB_TraceBuffer.st ---- *)
// Tampon circulaire de traces lu par la HMI depuis le dernier nSeq reçu (docs/05 § 9)
FUNCTION_BLOCK FB_TraceBuffer
VAR
    _refBuf : REFERENCE TO ST_TraceBuffer;
END_VAR

METHOD Bind
VAR_INPUT
    refBuf : REFERENCE TO ST_TraceBuffer;
END_VAR
_refBuf REF= refBuf;
END_METHOD

METHOD Add : UDINT
VAR_INPUT
    stTrace : ST_TraceRecord;
END_VAR
VAR
    k : INT;
END_VAR
IF NOT __ISVALIDREF(_refBuf) THEN RETURN; END_IF
_refBuf.nWriteSeq := _refBuf.nWriteSeq + 1;
k := UDINT_TO_INT(_refBuf.nWriteSeq MOD INT_TO_UDINT(GVL_Const.TRACE_BUFFER));
_refBuf.aTrace[k] := stTrace;
_refBuf.aTrace[k].nSeq := _refBuf.nWriteSeq;
Add := _refBuf.nWriteSeq;
END_METHOD
END_FUNCTION_BLOCK
